Fanuc KAREL source: ko00095.KL

-- PROVISIONAL review KL for V1013-1; original PC SHA256 f0d025db368703b1ee3fadc5697241725b7a90e64ce3f942bc8fe8cfa5ea54bd
-- Incomplete behavior may be omitted. Consult companion uncertainty JSON. Do not deploy.
PROGRAM KO00095
%NOLOCKGROUP
BEGIN
  -- UNRESOLVED_PC offsets 5-12; opcodes 9D,23
  -- UNRESOLVED_PC offsets 17-69; opcodes 27,27,49,7E,AD,27,49,7E,AD,22,31,7E,4A
  -- UNRESOLVED_PC offsets 74-78; opcodes 7F
END KO00095
